(* IEC 61131-3 sources: plc-st-coding-agent/progress/evidence/full_r8_20261110b/native_evidence/codex_minimax-m27/self-medium-05/1, 1 file *)

(* ---- candidate.st ---- *)
FUNCTION_BLOCK FB
VAR_INPUT
    enable       : BOOL;
    resetBtn     : BOOL;
    scanSeconds  : LREAL;
    steamFlow    : LREAL;
    fuelFlow     : LREAL;
    steamTemp    : LREAL;
    steamPressure: LREAL;
END_VAR
VAR_OUTPUT
    qualified    : BOOL;
    dataFault    : BOOL;
    qualifiedTon : LREAL;
    fuelTon      : LREAL;
    revenue      : LREAL;
    cost         : LREAL;
    netProfit    : LREAL;
END_VAR
VAR
    prevResetBtn : BOOL := FALSE;
    resetRising  : BOOL := FALSE;
END_VAR

resetRising := resetBtn AND NOT prevResetBtn;

qualified := (steamTemp >= 447.0) AND (steamTemp <= 453.0)
             AND (steamPressure >= 3750.0) AND (steamPressure <= 3850.0);

dataFault := (scanSeconds <= 0.0) OR (scanSeconds > 10.0)
             OR (steamFlow < 0.0) OR (steamFlow > 90.0)
             OR (fuelFlow < 0.0) OR (fuelFlow > 6.0);

IF resetRising THEN
    qualifiedTon := 0.0;
    fuelTon      := 0.0;
ELSIF enable AND NOT dataFault THEN
    qualifiedTon := qualifiedTon + steamFlow * scanSeconds / 1000.0;
    fuelTon      := fuelTon      + fuelFlow    * scanSeconds / 1000.0;
END_IF;

revenue   := qualifiedTon * 280.0;
cost      := fuelTon      * 1500.0;
netProfit := revenue - cost;

prevResetBtn := resetBtn;
END_FUNCTION_BLOCK
